Staubli VAL3: hmiAlert.pgx

public program hmiAlert(string x_sMsg, string x_sMsgType)
  local string l_sMsg
begin
  switch sLanguage
    case "english"
      l_sMsg=sAlertEN[x_sMsg]
    break
    case "chinese"
      l_sMsg=sAlertCN[x_sMsg]
    break
  endSwitch
  //*************************************************************
  utCtn_Message.Common.sSource="Page_Container_Alert.html"
  utTxt_popUpMsg.Common.sValue=l_sMsg
  //*************************************************************
  switch x_sMsgType
    case "info"
      utTxt_popUpMsg.Appearance.sBackgroundColour="#7C95FF"
    break
    //
    case "warning"
      utTxt_popUpMsg.Appearance.sBackgroundColour="#EEFB45"
    break
    //
    case "confirm"
      utTxt_popUpMsg.Appearance.sBackgroundColour="#FFFFFF"
    break
    //
    default
      utTxt_popUpMsg.Appearance.sBackgroundColour="#ADADB2"
    break
  endSwitch
  //*************************************************************
  if taskStatus("HmiClose")!=-1
    taskKill("HmiClose")
  endIf
  if taskStatus("HmiClose")==-1
    taskCreate "HmiClose",100,hmiClose()
  endIf
end
